(* IEC 61131-3 sources: plcassist-cli/packages/volt-lsp-iec/test-corpus/awa-palletizer/Device/Plc Logic/Application/Library Manager/CmpIecVarAccess Implementation, 36 files *)

(* ---- SVN_INFO_FLAGS.gvl ---- *)
VAR_GLOBAL
	XINCOMPLETE : BOOL := FALSE;
	XMODIFIED : BOOL := TRUE;
	XSWITCHED : BOOL := FALSE;
	XCLEAN : BOOL := FALSE;
	XDISCONNECTED : BOOL := FALSE;
END_VAR

(* ---- SVN_INFO_LASTCHANGE.gvl ---- *)
VAR_GLOBAL
	DTLASTCHANGEUTC : DATE_AND_TIME := DATE_AND_TIME#2021-4-1-14:23:38;
	WSLASTCHANGELOCAL : WSTRING(44) := "2021-04-01 16:23:38 +0200 (Thu, 01 Apr 2021)";
	WSLASTCHANGEAUTHOR : WSTRING(8) := "b.schurr";
END_VAR

(* ---- SVN_INFO_REVISIONS.gvl ---- *)
VAR_GLOBAL
	LIMINREVISION : LINT := LINT#52494;
	LIMAXREVISION : LINT := LINT#52494;
END_VAR

(* ---- SVN_INFO_SUMMARY.gvl ---- *)
VAR_GLOBAL
	SVERSIONSUMMARY : STRING(6) := '52494M';
END_VAR

(* ---- SVN_INFO_SUMMARYW.gvl ---- *)
VAR_GLOBAL
	WSVERSIONSUMMARY : WSTRING(6) := "52494M";
END_VAR

(* ---- SVN_INFO_URI.gvl ---- *)
VAR_GLOBAL
	WURL : WSTRING(129) := "svn://server04/LibrariesV3Source/branches/V3.5.17.0/System/SysLibs/CmpIecVarAccess Implementation/CmpIecVarAccess Implementation/";
END_VAR

(* ---- IECVARACCBROWSEDOWN2.fun ---- *)
FUNCTION IECVARACCBROWSEDOWN2 : ICollections.IBaseTreeNode
VAR_INPUT
	HINTERFACE : SysTypes.RTS_IEC_HANDLE;
	HNODE : ICollections.IBaseTreeNode;
	PVARIABLEINFORMATION : POINTER TO IecVarAccess_Interfaces.VariableInformationStruct3;
	PRESULT : POINTER TO SysTypes.RTS_IEC_RESULT;
END_VAR
END_FUNCTION

(* ---- IECVARACCBROWSEGETNEXT2.fun ---- *)
FUNCTION IECVARACCBROWSEGETNEXT2 : ICollections.IBaseTreeNode
VAR_INPUT
	HINTERFACE : SysTypes.RTS_IEC_HANDLE;
	HNODE : ICollections.IBaseTreeNode;
	PVARIABLEINFORMATION : POINTER TO IecVarAccess_Interfaces.VariableInformationStruct3;
	PRESULT : POINTER TO SysTypes.RTS_IEC_RESULT;
END_VAR
END_FUNCTION

(* ---- IECVARACCBROWSERECURSIVE.fun ---- *)
FUNCTION IECVARACCBROWSERECURSIVE : SysTypes.RTS_IEC_RESULT
VAR_INPUT
	HINTERFACE : SysTypes.RTS_IEC_HANDLE;
	HNODE : ICollections.IBaseTreeNode;
	PVARIABLEINFORMATION : POINTER TO IecVarAccess_Interfaces.VariableInformationStruct3;
	PFBROWSECALLBACK : POINTER TO BYTE;
	PUSERPARAMETER : POINTER TO BYTE;
END_VAR
END_FUNCTION

(* ---- IECVARACCBROWSEUP2.fun ---- *)
FUNCTION IECVARACCBROWSEUP2 : ICollections.IBaseTreeNode
VAR_INPUT
	HINTERFACE : SysTypes.RTS_IEC_HANDLE;
	HNODE : ICollections.IBaseTreeNode;
	PVARIABLEINFORMATION : POINTER TO IecVarAccess_Interfaces.VariableInformationStruct3;
	PRESULT : POINTER TO SysTypes.RTS_IEC_RESULT;
END_VAR
END_FUNCTION

(* ---- IECVARACCEXITVARINFO.fun ---- *)
FUNCTION IECVARACCEXITVARINFO : SysTypes.RTS_IEC_RESULT
VAR_INPUT
	PVARIABLEINFORMATION : POINTER TO IecVarAccess_Interfaces.VariableInformationStruct3;
END_VAR
END_FUNCTION

(* ---- IECVARACCGETFIRSTINTERFACE.fun ---- *)
FUNCTION IECVARACCGETFIRSTINTERFACE : IIecVarAccess3
VAR_INPUT
	PRESULT : POINTER TO RTS_IEC_RESULT;
END_VAR
END_FUNCTION

(* ---- IECVARACCGETFIRSTINTERFACE2.fun ---- *)
FUNCTION IECVARACCGETFIRSTINTERFACE2 : IBase
VAR_INPUT
	PRESULT : POINTER TO RTS_IEC_RESULT;
END_VAR
END_FUNCTION

(* ---- IECVARACCGETNEXTINTERFACE.fun ---- *)
FUNCTION IECVARACCGETNEXTINTERFACE : IIecVarAccess3
VAR_INPUT
	PIPREV : IIecVarAccess3;
	PRESULT : POINTER TO RTS_IEC_RESULT;
END_VAR
END_FUNCTION

(* ---- IECVARACCGETNEXTINTERFACE2.fun ---- *)
FUNCTION IECVARACCGETNEXTINTERFACE2 : IBase
VAR_INPUT
	PIPREV : IBase;
	PRESULT : POINTER TO RTS_IEC_RESULT;
END_VAR
END_FUNCTION

(* ---- IECVARACCGETNODE4.fun ---- *)
FUNCTION IECVARACCGETNODE4 : ICollections.IBaseTreeNode
VAR_INPUT
	PSZPATH : POINTER TO STRING;
	PHINTERFACE : POINTER TO SysTypes.RTS_IEC_HANDLE;
	PVARIABLEINFORMATION : POINTER TO IecVarAccess_Interfaces.VariableInformationStruct3;
	PRESULT : POINTER TO SysTypes.RTS_IEC_RESULT;
END_VAR
END_FUNCTION

(* ---- IECVARACCGETNODEFULLPATH4.fun ---- *)
FUNCTION IECVARACCGETNODEFULLPATH4 : DINT
VAR_INPUT
	HINTERFACE : SysTypes.RTS_IEC_HANDLE;
	HNODE : ICollections.IBaseTreeNode;
	PVARIABLEINFORMATION : POINTER TO IecVarAccess_Interfaces.VariableInformationStruct3;
	PSZPATH : POINTER TO STRING;
	IMAXPATH : DINT;
	PRESULT : POINTER TO SysTypes.RTS_IEC_RESULT;
END_VAR
END_FUNCTION

(* ---- IECVARACCGETNODENAME4.fun ---- *)
FUNCTION IECVARACCGETNODENAME4 : SysTypes.RTS_IEC_RESULT
VAR_INPUT
	HINTERFACE : SysTypes.RTS_IEC_HANDLE;
	HNODE : ICollections.IBaseTreeNode;
	PVARIABLEINFORMATION : POINTER TO IecVarAccess_Interfaces.VariableInformationStruct3;
	PSZNODENAME : POINTER TO STRING;
	NNODENAMELEN : UDINT;
END_VAR
END_FUNCTION

(* ---- IECVARACCGETSYMBOLSETMASK.fun ---- *)
FUNCTION IECVARACCGETSYMBOLSETMASK : DWORD
VAR_INPUT
	HUSER : RTS_IEC_HANDLE;
	HINTERFACE : RTS_IEC_HANDLE;
	PRESULT : POINTER TO RTS_IEC_RESULT;
END_VAR
END_FUNCTION

(* ---- IECVARACCINITVARINFO.fun ---- *)
FUNCTION IECVARACCINITVARINFO : SysTypes.RTS_IEC_RESULT
VAR_INPUT
	PVARIABLEINFORMATION : POINTER TO IecVarAccess_Interfaces.VariableInformationStruct3;
	NSIZEOFVARINFO : UINT;
END_VAR
END_FUNCTION

(* ---- IECVARACCINITVARINFO2.fun ---- *)
FUNCTION IECVARACCINITVARINFO2 : SysTypes.RTS_IEC_RESULT
VAR_INPUT
	PVARIABLEINFORMATION : POINTER TO IecVarAccess_Interfaces.VariableInformationStruct3;
	NSIZEOFVARINFO : UINT;
	HUSER : RTS_IEC_HANDLE;
END_VAR
END_FUNCTION

(* ---- IECVARACCINVALIDATENODE.fun ---- *)
FUNCTION IECVARACCINVALIDATENODE : RTS_IEC_RESULT
VAR_INPUT
	HNODE : RTS_IEC_HANDLE;
END_VAR
END_FUNCTION

(* ---- IECVARACCNODEINFOADDBROWSEINFO.fun ---- *)
FUNCTION IECVARACCNODEINFOADDBROWSEINFO : SysTypes.RTS_IEC_RESULT
VAR_INPUT
	PVARIABLEINFORMATION : POINTER TO IecVarAccess_Interfaces.VariableInformationStruct3;
	PBROWSEINFODATA : POINTER TO RtsBrowseInfo;
END_VAR
END_FUNCTION

(* ---- IECVARACCNODEINFOADDREFERENCE.fun ---- *)
FUNCTION IECVARACCNODEINFOADDREFERENCE : SysTypes.RTS_IEC_RESULT
VAR_INPUT
	PVARIABLEINFORMATION : POINTER TO IecVarAccess_Interfaces.VariableInformationStruct3;
	PREFERENCEINFODATA : POINTER TO BYTE;
	NINFOSIZE : XWORD;
	PNEWREFERENCEINFO : POINTER TO POINTER TO BYTE;
END_VAR
END_FUNCTION

(* ---- IECVARACCNODEINFOGETBROWSEINFO.fun ---- *)
FUNCTION IECVARACCNODEINFOGETBROWSEINFO : POINTER TO RtsBrowseInfo
VAR_INPUT
	PVARIABLEINFORMATION : POINTER TO IecVarAccess_Interfaces.VariableInformationStruct3;
	PLAST : POINTER TO RtsBrowseInfo;
	PRESULT : POINTER TO SysTypes.RTS_IEC_RESULT;
END_VAR
END_FUNCTION

(* ---- IECVARACCNODEINFOGETREFERENCE.fun ---- *)
FUNCTION IECVARACCNODEINFOGETREFERENCE : POINTER TO BYTE
VAR_INPUT
	PVARIABLEINFORMATION : POINTER TO IecVarAccess_Interfaces.VariableInformationStruct3;
	PRESULT : POINTER TO SysTypes.RTS_IEC_RESULT;
END_VAR
END_FUNCTION

(* ---- IECVARACCNODEINFOREMOVEBROWSEINFO.fun ---- *)
FUNCTION IECVARACCNODEINFOREMOVEBROWSEINFO : SysTypes.RTS_IEC_RESULT
VAR_INPUT
	PVARIABLEINFORMATION : POINTER TO IecVarAccess_Interfaces.VariableInformationStruct3;
END_VAR
END_FUNCTION

(* ---- IECVARACCNODEINFOREMOVEREFERENCE.fun ---- *)
FUNCTION IECVARACCNODEINFOREMOVEREFERENCE : SysTypes.RTS_IEC_RESULT
VAR_INPUT
	PVARIABLEINFORMATION : POINTER TO IecVarAccess_Interfaces.VariableInformationStruct3;
END_VAR
END_FUNCTION

(* ---- IECVARACCREGISTERINSTANCE.fun ---- *)
FUNCTION IECVARACCREGISTERINSTANCE : RTS_IEC_HANDLE
VAR_INPUT
	PIIECVARACCESS : CmpIecVarAccess_Interfaces.IIecVarAccess;
	PRESULT : POINTER TO RTS_IEC_RESULT;
END_VAR
END_FUNCTION

(* ---- IECVARACCREGISTERINSTANCE2.fun ---- *)
FUNCTION IECVARACCREGISTERINSTANCE2 : RTS_IEC_HANDLE
VAR_INPUT
	PIIECVARACCESS2 : CmpIecVarAccess_Interfaces.IIecVarAccess2;
	PRESULT : POINTER TO RTS_IEC_RESULT;
END_VAR
END_FUNCTION

(* ---- IECVARACCREGISTERINSTANCE3.fun ---- *)
FUNCTION IECVARACCREGISTERINSTANCE3 : RTS_IEC_HANDLE
VAR_INPUT
	PIIECVARACCESS3 : IIecVarAccess3;
	PRESULT : POINTER TO RTS_IEC_RESULT;
END_VAR
END_FUNCTION

(* ---- IECVARACCREGISTERINSTANCEBASE.fun ---- *)
FUNCTION IECVARACCREGISTERINSTANCEBASE : RTS_IEC_HANDLE
VAR_INPUT
	PIBASE : IBase;
	PRESULT : POINTER TO RTS_IEC_RESULT;
END_VAR
END_FUNCTION

(* ---- IECVARACCREGISTERINSTANCEBASE2.fun ---- *)
FUNCTION IECVARACCREGISTERINSTANCEBASE2 : RTS_IEC_HANDLE
VAR_INPUT
	PIBASE : IBase;
	UDICRC : UDINT;
	PRESULT : POINTER TO RTS_IEC_RESULT;
END_VAR
END_FUNCTION

(* ---- IECVARACCSETSYMBOLCONFIGCRC.fun ---- *)
FUNCTION IECVARACCSETSYMBOLCONFIGCRC : RTS_IEC_RESULT
VAR_INPUT
	HINSTANCE : RTS_IEC_HANDLE;
	UDICRC : UDINT;
END_VAR
END_FUNCTION

(* ---- IECVARACCUNREGISTERINSTANCE.fun ---- *)
FUNCTION IECVARACCUNREGISTERINSTANCE : RTS_IEC_RESULT
VAR_INPUT
	HINSTANCE : RTS_IEC_HANDLE;
END_VAR
END_FUNCTION

(* ---- IECVARACCUPDATESYMBOLSETS.fun ---- *)
FUNCTION IECVARACCUPDATESYMBOLSETS : RTS_IEC_RESULT
VAR_INPUT
	HINTERFACE : RTS_IEC_HANDLE;
	PSYMBOLSSETS : POINTER TO IecVarAccSymbolSetDescription;
	NUMOFSYMBOLSSETS : UDINT;
END_VAR
END_FUNCTION
